// TIA Portal V21 export
FUNCTION_BLOCK "FB_PumpInterlockLad"   // FB110, LAD
TITLE = Блокировки насоса по уровню и давлению (LAD)
{ S7_Optimized_Access := 'TRUE' }
AUTHOR : WTP2
FAMILY : Drives
VERSION : 0.1
// Блокировки насоса II подъёма по уровню в РЧВ и давлению в коллекторе (LAD).
// 1. xLowLevel := iLevel_cm < iLevelMin_cm.  2. xHighPress := iPressure_kPa > iPressureMax_kPa.
// 3. Если xLowLevel OR xHighPress — установить xAlarmLatch (S).
// 4. Если xAck AND NOT xLowLevel AND NOT xHighPress — сбросить xAlarmLatch (R).
// 5. Обслуживание: при xMaint прыжок вперёд к метке NoAuto (сети 6-7 не выполняются).
// 6. xPumpOn := xAutoReq AND NOT xAlarmLatch.
// 7. По фронту xPumpOn (P_TRIG, бит xRunEdge): iRunCount := iRunCount + 1 (ADD Int); xCountOk := ENO сложения
//    (ENO = 0 при переполнении Int: 32767 + 1).
// 8. Метка NoAuto: при xMaint сбросить xPumpOn (R).
// 9. При xPumpOn — цепочка трёх вызовов FC_ClampPctLad через EN/ENO: iStage1 := clamp(iLevel_cm, 0, 100);
//    iStage2 := clamp(iStage1, 10, 90); iSetpoint_pct := clamp(iStage2, 20, 80); xChainOk := ENO третьего вызова.
// 10. При NOT xPumpOn: iSetpoint_pct := 0 (MOVE).
// 11. xAlarm := xAlarmLatch.  12. xRunMem := xRunEdge (бит памяти фронта читается в другой сети).
// stored: AutoNumber false, SetENOAutomatically false
   VAR_INPUT
      xAutoReq : Bool;   // Запрос автоматики на работу
      iLevel_cm : Int;   // Уровень в РЧВ, см
      iLevelMin_cm : Int := 50;   // Минимальный уровень, см
      iPressure_kPa : Int;   // Давление в коллекторе, кПа
      iPressureMax_kPa : Int := 600;   // Максимальное давление, кПа
      xAck : Bool;   // Квитирование аварии
      xMaint : Bool;   // Режим обслуживания
   END_VAR
   VAR_OUTPUT
      xPumpOn : Bool;   // Команда насосу
      xLowLevel : Bool;   // Низкий уровень
      xHighPress : Bool;   // Высокое давление
      xAlarm : Bool;   // Авария (защёлка)
      iRunCount : Int;   // Число включений
      xCountOk : Bool;   // ENO сложения: нет переполнения
      iSetpoint_pct : Int;   // Уставка производительности, %
      xChainOk : Bool;   // ENO цепочки вызовов
      xRunMem : Bool;   // Копия бита памяти фронта
   END_VAR
   VAR
      xAlarmLatch : Bool;   // Защёлка аварии
      xRunEdge : Bool;   // Бит памяти фронта xPumpOn
      iStage1 : Int;   // Уставка после первого ограничения
      iStage2 : Int;   // Уставка после второго ограничения
   END_VAR
   VAR_TEMP   // added for the SCL form of the ladder/FBD networks
      _w1 : Bool;
      _w2 : Bool;
      _w3 : Bool;
   END_VAR
BEGIN

REGION Network 1: Низкий уровень в РЧВ
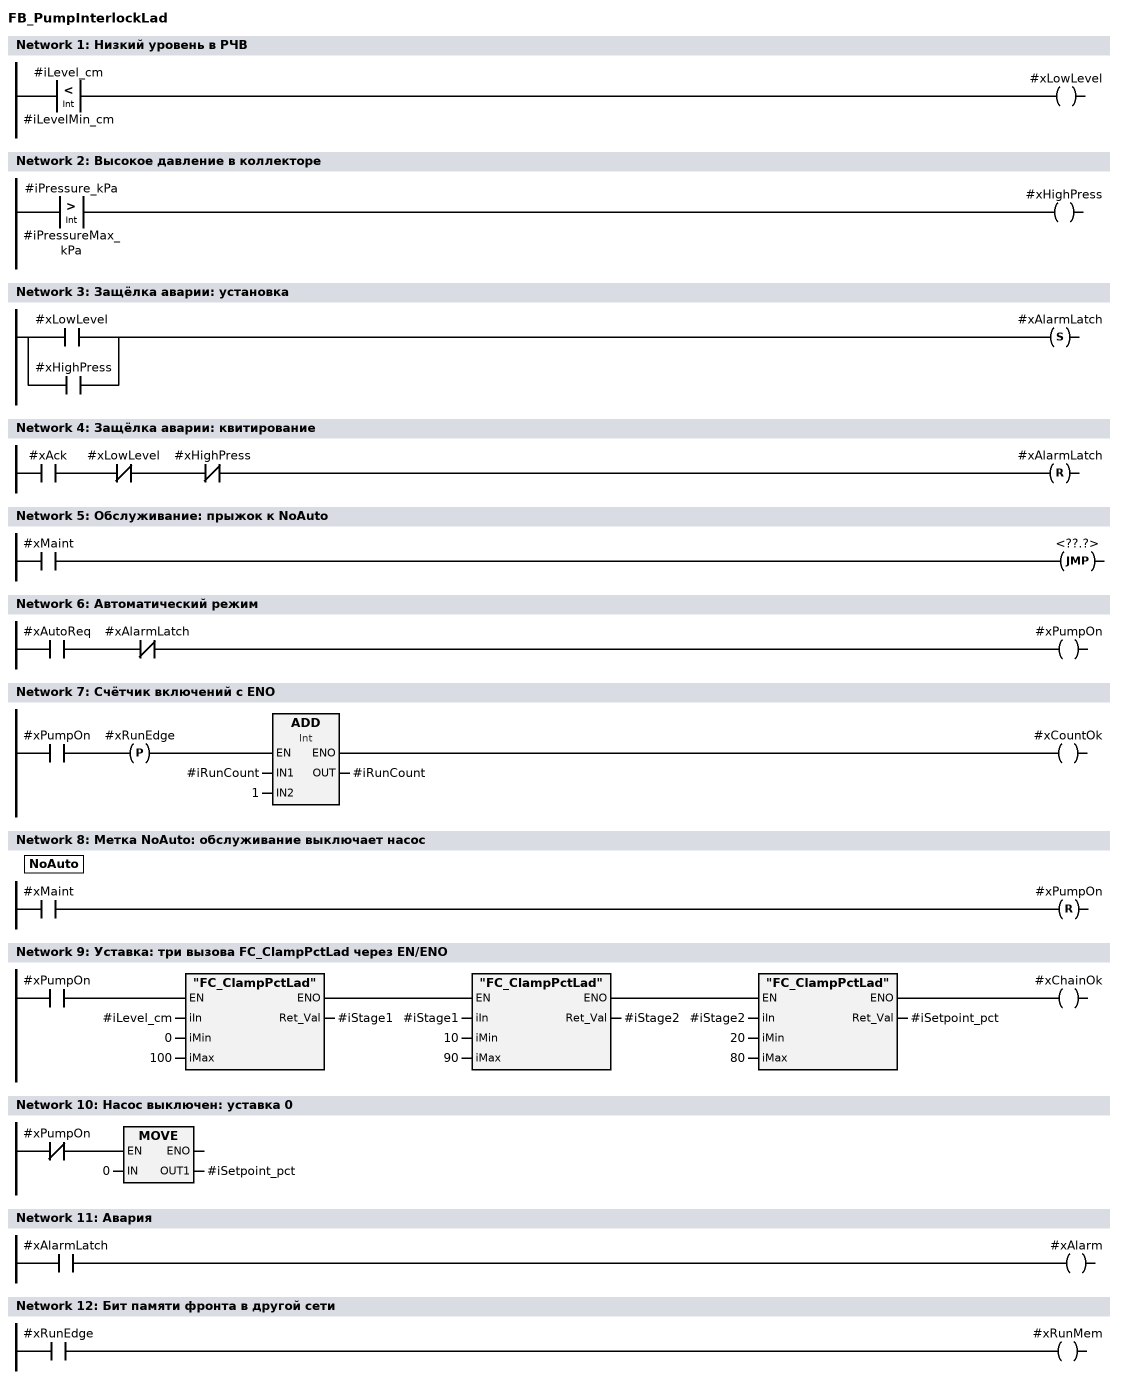
   RUNG wire#powerrail
      { S7_Templates := "SrcType := Int" } LT_Contact(in1 := #iLevel_cm, in2 := #iLevelMin_cm)
      Coil( #xLowLevel )
   END_RUNG
   // the same network as SCL:
   #xLowLevel := #iLevel_cm < #iLevelMin_cm;
END_REGION

REGION Network 2: Высокое давление в коллекторе
   RUNG wire#powerrail
      { S7_Templates := "SrcType := Int" } GT_Contact(in1 := #iPressure_kPa, in2 := #iPressureMax_kPa)
      Coil( #xHighPress )
   END_RUNG
   // the same network as SCL:
   #xHighPress := #iPressure_kPa > #iPressureMax_kPa;
END_REGION

REGION Network 3: Защёлка аварии: установка
   RUNG wire#powerrail
      Contact( #xLowLevel )
      wire#w1
      S_Coil( #xAlarmLatch )
   END_RUNG
   RUNG wire#powerrail
      Contact( #xHighPress )
   END_RUNG wire#w1
   // the same network as SCL:
   IF #xLowLevel OR #xHighPress THEN #xAlarmLatch := TRUE; END_IF;
END_REGION

REGION Network 4: Защёлка аварии: квитирование
   RUNG wire#powerrail
      Contact( #xAck )
      I_Contact( #xLowLevel )
      I_Contact( #xHighPress )
      R_Coil( #xAlarmLatch )
   END_RUNG
   // the same network as SCL:
   IF #xAck AND NOT #xLowLevel AND NOT #xHighPress THEN #xAlarmLatch := FALSE; END_IF;
END_REGION

REGION Network 5: Обслуживание: прыжок к NoAuto
   IF #xMaint THEN GOTO <??.?>; END_IF;
END_REGION

REGION Network 6: Автоматический режим
   RUNG wire#powerrail
      Contact( #xAutoReq )
      I_Contact( #xAlarmLatch )
      Coil( #xPumpOn )
   END_RUNG
   // the same network as SCL:
   #xPumpOn := #xAutoReq AND NOT #xAlarmLatch;
END_REGION

REGION Network 7: Счётчик включений с ENO
   // ENO of a box is taken as its EN; it also drops when the box reports an error
   #_w1 := #xPumpOn AND NOT #xRunEdge;   // rising edge
   #xRunEdge := #xPumpOn;
   IF #_w1 THEN #iRunCount := #iRunCount + 1; END_IF;
   #xCountOk := #_w1;
END_REGION

REGION Network 8: Метка NoAuto: обслуживание выключает насос
   Label( NoAuto )
   RUNG wire#powerrail
      Contact( #xMaint )
      R_Coil( #xPumpOn )
   END_RUNG
   // the same network as SCL:
   NoAuto:
   IF #xMaint THEN #xPumpOn := FALSE; END_IF;
END_REGION

REGION Network 9: Уставка: три вызова FC_ClampPctLad через EN/ENO
   RUNG wire#powerrail
      Contact( #xPumpOn )
      "FC_ClampPctLad"(iIn := #iLevel_cm, iMin := 0, iMax := 100, Ret_Val => #iStage1)
      "FC_ClampPctLad"(iIn := #iStage1, iMin := 10, iMax := 90, Ret_Val => #iStage2)
      "FC_ClampPctLad"(iIn := #iStage2, iMin := 20, iMax := 80, Ret_Val => #iSetpoint_pct)
      Coil( #xChainOk )
   END_RUNG
   // the same network as SCL:
   #iStage1 := "FC_ClampPctLad"(EN := #xPumpOn, iIn := #iLevel_cm, iMin := 0, iMax := 100, ENO => #_w1);
   #iStage2 := "FC_ClampPctLad"(EN := #_w1, iIn := #iStage1, iMin := 10, iMax := 90, ENO => #_w2);
   #iSetpoint_pct := "FC_ClampPctLad"(EN := #_w2, iIn := #iStage2, iMin := 20, iMax := 80, ENO => #_w3);
   #xChainOk := #_w3;
END_REGION

REGION Network 10: Насос выключен: уставка 0
   IF NOT #xPumpOn THEN #iSetpoint_pct := 0; END_IF;
END_REGION

REGION Network 11: Авария
   RUNG wire#powerrail
      Contact( #xAlarmLatch )
      Coil( #xAlarm )
   END_RUNG
   // the same network as SCL:
   #xAlarm := #xAlarmLatch;
END_REGION

REGION Network 12: Бит памяти фронта в другой сети
   RUNG wire#powerrail
      Contact( #xRunEdge )
      Coil( #xRunMem )
   END_RUNG
   // the same network as SCL:
   #xRunMem := #xRunEdge;
END_REGION
END_FUNCTION_BLOCK
